TYPE ST_Recipe :
STRUCT
	fLevelSetpoint : REAL := 80.0;   // fill level to reach in %
	tSettle : TIME := T#5S;          // how long the product settles
	(* recipe number from MES *)
	nRecipeNo : DINT;
	sName : STRING(40);
END_STRUCT
END_TYPE

(* stored: Version 1.1.0.1, ProductVersion 3.1.4026.12
   DUT ST_Recipe: Id {1a2b3c4d-0000-4000-8000-000000000002} *)
